Universal Robots URScript: T009_zai-org_GLM-4.7-FP8_edit_perf_rep1.urscript

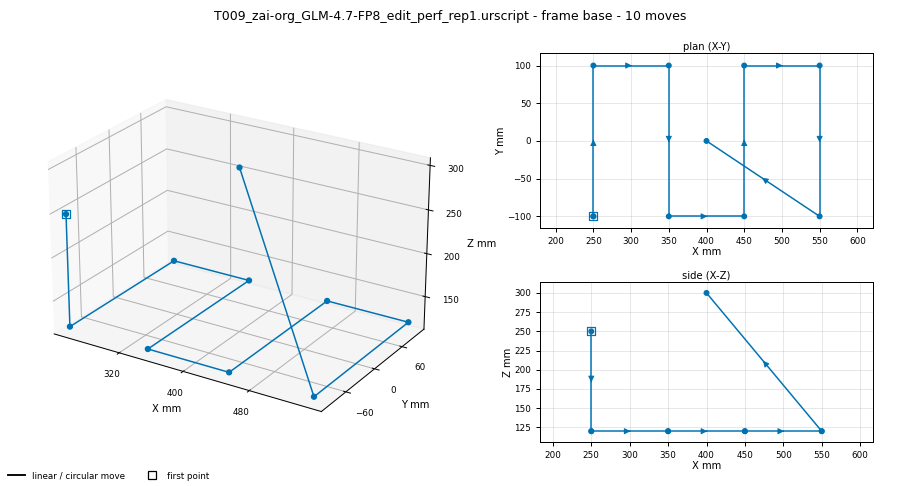
[picture p0: tool path of T009_zai-org_GLM-4.7-FP8_edit_perf_rep1.urscript in frame base, 10 of 12 moves have a stored position in this frame; points joined in program order, loops and branches not executed]
# Task: T009 — Laser surface scan — fenced mode (OPTIMIZED)
# Optimized for reduced cycle time
# Operating mode: fenced | Max TCP speed: 0.200 m/s
# Robot: ur5e
#
# WARNING: This is auto-generated code for SIMULATION ONLY.
# Do NOT deploy to a physical robot without safety review.

def task_T009():
  # [0] Home - Increased joint velocity and acceleration for faster transit
  movej([0.0000, -1.5708, 1.5708, -1.5708, -1.5708, 0.0000], a=3.0000, v=2.5000)

  # [1] Above scan start - Max speed, increased acceleration
  movel(p[0.250000, -0.100000, 0.250000, 0.0000, 3.1416, 0.0000], a=1.2000, v=0.2000, r=0.0100)

  # [2] Descend to scan height - Max speed, increased acceleration
  movel(p[0.250000, -0.100000, 0.120000, 0.0000, 3.1416, 0.0000], a=1.2000, v=0.2000, r=0.0100)

  # [3] Laser ON
  set_digital_out(3, True)

  # [4] Scan line 1 - Max speed, increased acceleration
  movel(p[0.250000, 0.100000, 0.120000, 0.0000, 3.1416, 0.0000], a=1.2000, v=0.2000, r=0.0100)

  # [5] Step to line 2 - Max speed, increased acceleration
  movel(p[0.350000, 0.100000, 0.120000, 0.0000, 3.1416, 0.0000], a=1.2000, v=0.2000, r=0.0100)

  # [6] Scan line 2 reverse - Max speed, increased acceleration
  movel(p[0.350000, -0.100000, 0.120000, 0.0000, 3.1416, 0.0000], a=1.2000, v=0.2000, r=0.0100)

  # [7] Step to line 3 - Max speed, increased acceleration
  movel(p[0.450000, -0.100000, 0.120000, 0.0000, 3.1416, 0.0000], a=1.2000, v=0.2000, r=0.0100)

  # [8] Scan line 3 - Max speed, increased acceleration
  movel(p[0.450000, 0.100000, 0.120000, 0.0000, 3.1416, 0.0000], a=1.2000, v=0.2000, r=0.0100)

  # [9] Step to line 4 - Max speed, increased acceleration
  movel(p[0.550000, 0.100000, 0.120000, 0.0000, 3.1416, 0.0000], a=1.2000, v=0.2000, r=0.0100)

  # [10] Scan line 4 reverse - Max speed, increased acceleration, stop at end
  movel(p[0.550000, -0.100000, 0.120000, 0.0000, 3.1416, 0.0000], a=1.2000, v=0.2000, r=0.0)

  # [11] Laser OFF
  set_digital_out(3, False)

  # [12] Retract - Max speed, increased acceleration
  movel(p[0.400000, 0.000000, 0.300000, 0.0000, 3.1416, 0.0000], a=1.2000, v=0.2000, r=0.0100)

  # [13] Return home - Increased joint velocity and acceleration
  movej([0.0000, -1.5708, 1.5708, -1.5708, -1.5708, 0.0000], a=3.0000, v=2.5000)

end

# Entry point
task_T009()
